// TIA Portal V20 export
// export: Created 2026-10-12T16:46:22.1158702Z, ExportSetting WithDefaults, DisplayName Totally Integrated Automation Portal, DisplayVersion V20 Update 6, DisplayName TIA Portal Openness, DisplayVersion V20 Update 6, DisplayName TIA Portal Version Control Interface, DisplayVersion V20 Update 6, DisplayName SINAMICS Startdrive Advanced, DisplayVersion V20 SP1 Update 2, DisplayName SINAMICS Startdrive G110M, G120, G120C, G120D, G120P, G115D, DisplayVersion V20 SP1 Update 2, DisplayName SINAMICS Startdrive G130, G150, S120, S150, SINAMICS MV, G220, S200, S210, DisplayVersion V20 SP1 Update 2, DisplayName STEP 7 Professional, DisplayVersion V20 Update 6, DisplayName STEP 7 Safety, DisplayVersion V20 Update 2, DisplayName WinCC Basic/Comfort/Advanced, DisplayVersion V20 Update 6, DisplayName WinCC Professional, DisplayVersion V20 Update 6, DisplayName WinCC Unified, DisplayVersion V20 Update 6
VAR_GLOBAL   // PLC tag table "Standard-Variablentabelle"
   "FI-Schutz 200F1 Heizung Bad 7 ist O.K." AT %I2.2 : Bool;
   "Sicherheitsschuetz Rueckfuehrung Heizung Bad 7" AT %I2.3 : Bool;
   "Heizung Bad 7 Keine uebertemperatur" AT %I2.4 : Bool;
   "Störmeldung Ultraschall Bad 7" AT %I2.6 : Bool;
   "Niveau Bad 7 OK" AT %I10.0 : Bool;
   "Pt100 Heizung Bad 7" AT %IW60 : Word;
   "FI-Schutz 210F1 Heizung Bad 8 ist O.K." AT %I2.7 : Bool;
   "Sicherheitsschuetz Rueckfuehrung Heizung Bad 8" AT %I3.0 : Bool;
   "Heizung Bad 8 Keine uebertemperatur" AT %I3.1 : Bool;
   "FILS Automat 213F1 Ultraschall Bad 8 ist O.K." AT %I3.2 : Bool;
   "Störmeldung Ultraschall Bad 8" AT %I3.3 : Bool;
   "Motorschutz 215Q1 Pumpe Bad 8 ist O.K." AT %I3.4 : Bool;
   "Wartungsschalter Pumpe Bad 8 ist eingeschaltet" AT %I3.5 : Bool;
   "Niveau Bad 8 OK" AT %I10.1 : Bool;
   "FI-Schutz 220F1 Heizung Bad 12 ist O.K." AT %I3.6 : Bool;
   "Sicherheitsschuetz Rueckfuehrung Heizung Bad 12" AT %I3.7 : Bool;
   "Heizung Bad 12 Keine uebertemperatur" AT %I4.0 : Bool;
   "FILS Automat 223F1 Ultraschall Bad 12 ist O.K." AT %I4.1 : Bool;
   "Störmeldung Ultraschall Bad 12" AT %I4.2 : Bool;
   "Motorschutz 225Q1 Pumpe Bad 12 ist O.K." AT %I4.3 : Bool;
   "Wartungsschalter Pumpe Bad 12 ist eingeschaltet" AT %I4.4 : Bool;
   "Niveau Bad 12 OK" AT %I10.2 : Bool;
   "Motorschutz 235Q1 Pumpe Bad 14 ist O.K." AT %I4.5 : Bool;
   "Wartungsschalter Pumpe Bad 14 ist eingeschaltet" AT %I4.6 : Bool;
   "Motorschutz 245Q1 Pumpe Bad 18 ist O.K." AT %I4.7 : Bool;
   "Wartungsschalter Pumpe Bad 18 ist eingeschaltet" AT %I5.0 : Bool;
   "Motorschutz 255Q1 Pumpe Bad 19 ist O.K." AT %I5.1 : Bool;
   "Wartungsschalter Pumpe Bad 19 ist eingeschaltet" AT %I5.2 : Bool;
   "Motorschutz 265Q1 Pumpe Bad 21 ist O.K." AT %I5.3 : Bool;
   "Wartungsschalter Pumpe Bad 21 ist eingeschaltet" AT %I5.4 : Bool;
   "Motorschutz und FI-Schutz 270Q1, 270F1 Heizung Bad 25 sind O.K." AT %I5.5 : Bool;
   "Motorschutz und FI-Schutz 271Q1, 271F1 Heizung Bad 25 sind O.K." AT %I5.6 : Bool;
   "Sicherheitsschuetze Rueckfuehrung Heizung Bad 25" AT %I5.7 : Bool;
   "Heizung Bad 25 Keine uebertemperatur" AT %I6.0 : Bool;
   "FILS Automat 274F1 Analysegerät Bad 25 ist O.K." AT %I6.1 : Bool;
   "Motorschutz 275Q1 Pumpe Bad 25 ist O.K." AT %I6.2 : Bool;
   "Wartungsschalter Pumpe Bad 25 ist eingeschaltet" AT %I6.3 : Bool;
   "Motorschutz 276Q1 Warenbewegung 1 Bad 25 ist O.K." AT %I6.4 : Bool;
   "Motorschutz 277Q1 Warenbewegung 2 Bad 25 ist O.K." AT %I6.5 : Bool;
   "FILS Automat 203F1 GR Wannenschutz Bad 25 ist O.K." AT %I2.5 : Bool;
   "Motorschutz 275aQ1 Pumpe Bad 25 ist O.K." AT %I8.7 : Bool;
   "Warenbewegung 1 Bad 25 FU bereit" AT %I9.5 : Bool;
   "Warenbewegung 2 Bad 25 FU bereit" AT %I9.6 : Bool;
   "Wartungsschalter Pumpe Bad 25 ist eingeschaltet(1)" AT %I9.7 : Bool;
   "Niveau Bad 25 OK" AT %I10.3 : Bool;
   "Motorschutz 285Q1 Pumpe Bad 26 ist O.K." AT %I6.6 : Bool;
   "Wartungsschalter Pumpe Bad 26 ist eingeschaltet" AT %I6.7 : Bool;
   "Motorschutz 295Q1 Pumpe Bad 31 ist O.K." AT %I7.0 : Bool;
   "Wartungsschalter Pumpe Bad 31 ist eingeschaltet" AT %I7.1 : Bool;
   "FI-Schutz 300F1 Heizung Bad 36 ist O.K." AT %I7.2 : Bool;
   "Sicherheitsschuetz Rueckfuehrung Heizung Bad 36" AT %I7.3 : Bool;
   "Heizung Bad 36 Keine uebertemperatur" AT %I7.4 : Bool;
   "Niveau Bad 36 OK" AT %I10.4 : Bool;
   "FI-Schutz 310F1 Heizung Bad 40 ist O.K." AT %I7.5 : Bool;
   "Sicherheitsschuetz Rueckfuehrung Heizung Bad 40" AT %I7.6 : Bool;
   "Heizung Bad 40 Keine uebertemperatur" AT %I7.7 : Bool;
   "Motorschutz 325Q1 Pumpe Bad 41 ist O.K." AT %I8.0 : Bool;
   "Wartungsschalter Pumpe Bad 41 ist eingeschaltet" AT %I8.1 : Bool;
   "Motorschutz 335Q1 Pumpe Bad 45 ist O.K." AT %I8.2 : Bool;
   "Wartungsschalter Pumpe Bad 45 ist eingeschaltet" AT %I8.3 : Bool;
   "FI-Schutz 340F1 Heizung Bad 46 ist O.K." AT %I8.4 : Bool;
   "Sicherheitsschuetz Rueckfuehrung Heizung Bad 46" AT %I8.5 : Bool;
   "Heizung Bad 46 Keine uebertemperatur" AT %I8.6 : Bool;
   "Niveau Bad 46 OK" AT %I10.6 : Bool;
   "Motorschutz 15Q0 Schaltschrankklimatisierung Feld 1-4 ist O.K." AT %I0.0 : Bool;
   "Klimagerät +E1-15A0 ist in Ordnung" AT %I0.1 : Bool;
   "Schaltschranktemperatur Feld 1 ist zu hoch" AT %I0.2 : Bool;
   "Schaltschranktemperatur Feld 2 ist zu hoch" AT %I0.3 : Bool;
   "FILS Automat 19F1 Schuko.Steckdosen PC-Bildschirm ist O.K." AT %I0.4 : Bool;
   "Not-Aus ist OK" AT %I0.5 : Bool;
   "Steuerspannung 31F1 Schaltschrank E1 ist O.K." AT %I1.0 : Bool;
   "Steuerspannung 31F3 SPS Out 1 ist O.K." AT %I1.1 : Bool;
   "Steuerspannung 31F5 SPS Out 2 ist O.K." AT %I1.2 : Bool;
   "Steuerspannung 31F6 SPS Out 3 ist O.K." AT %I1.3 : Bool;
   "Steuerspannung 31F8 Out 4 ist O.K." AT %I1.4 : Bool;
   "Steuerspannung 32F1 Rueckmeldung Wartungsschalter ist O.K." AT %I1.5 : Bool;
   "Steuerspannung 32F3 Sensorik 1 ist O.K." AT %I1.6 : Bool;
   "Busspannung 41F1 ist ok" AT %I1.7 : Bool;
   "Busspannung 41F2 ist ok" AT %I2.0 : Bool;
   "Busspannung 41F4 ist ok" AT %I2.1 : Bool;
   "Pt100 Heizung Bad 8" AT %IW62 : Word;
   "Pt100 Heizung Bad 12" AT %IW64 : Word;
   "Pt100 Heizung Bad 25" AT %IW66 : Word;
   "Pt100 Heizung Bad 36" AT %IW68 : Word;
   "Pt100 Heizung Bad 40" AT %IW70 : Word;
   "Pt100 Heizung Bad 46" AT %IW72 : Word;
   "FU Pumpe bereit" AT %I0.7 : Bool;
   Flexkraft_1 AT %IW500 : Word;
   Flexkraft_2 AT %IW502 : Word;
   Flexkraft_3 AT %IW504 : Word;
   Flexkraft_4 AT %IW506 : Word;
   Flexkraft_5 AT %IW508 : Word;
   Flexkraft_6 AT %IW510 : Word;
   Flexkraft_7 AT %IW512 : Word;
   Flexkraft_8 AT %IW514 : Word;
   Flexkraft_9 AT %IW516 : Word;
   Flexkraft_10 AT %IW518 : Word;
   "Niveau Bad 40 OK" AT %I10.5 : Bool;
   "Regelung Heizung Bad 7" AT %Q2.0 : Bool;
   "Sicherheitsschuetz Heizung Bad 7" AT %Q2.1 : Bool;
   "Pumpe Bad 8" AT %Q0.0 : Bool;
   "Regelung Heizung Bad 8" AT %Q2.2 : Bool;
   "Sicherheitsschuetz Heizung Bad 8" AT %Q2.3 : Bool;
   "Pumpe Bad 12" AT %Q0.1 : Bool;
   "Regelung Heizung Bad 12" AT %Q2.4 : Bool;
   "Sicherheitsschuetz Heizung Bad 12" AT %Q2.5 : Bool;
   "Pumpe Bad 14" AT %Q0.2 : Bool;
   "Pumpe Bad 18" AT %Q0.3 : Bool;
   "Pumpe Bad 19" AT %Q0.4 : Bool;
   "Pumpe Bad 21" AT %Q0.5 : Bool;
   "Netzschuetz Pumpe Bad 25" AT %Q0.6 : Bool;
   "Warenbewegung 1 Bad 25 Freigabe FU" AT %Q1.3 : Bool;
   "Warenbewegung 1 Bad 25 Reset FU" AT %Q1.4 : Bool;
   "Warenbewegung 2 Bad 25 Freigabe FU" AT %Q1.5 : Bool;
   "Warenbewegung 2 Bad 25 Reset FU" AT %Q1.6 : Bool;
   "Ansteuerung 275aK8" AT %Q1.7 : Bool;
   "Regelung Heizung 1 Bad 25" AT %Q2.6 : Bool;
   "Regelung Heizung 2 Bad 25" AT %Q2.7 : Bool;
   "Sicherheitsschuetze Heizung 1 + 2 Bad 25" AT %Q3.0 : Bool;
   "Warenbewegung 1 Bad 25 Netzschuetz" AT %Q3.1 : Bool;
   "Warenbewegung 2 Bad 25 Netzschuetz" AT %Q3.2 : Bool;
   "Pumpe Bad 26" AT %Q0.7 : Bool;
   "Pumpe Bad 31" AT %Q1.0 : Bool;
   "Regelung Heizung Bad 36" AT %Q3.3 : Bool;
   "Sicherheitsschuetz Heizung Bad 36" AT %Q3.4 : Bool;
   "Regelung Heizung Bad 40" AT %Q3.5 : Bool;
   "Sicherheitsschuetz Heizung Bad 40" AT %Q3.6 : Bool;
   "Pumpe Bad 41" AT %Q1.1 : Bool;
   "Pumpe Bad 45" AT %Q1.2 : Bool;
   "Regelung Heizung Bad 46" AT %Q3.7 : Bool;
   "Sicherheitsschuetz Heizung Bad 46" AT %Q4.0 : Bool;
   "Masch.Leuchte 1 Anlage Hupe" AT %Q4.1 : Bool;
   "Freigabe Ultraschall Pos. 8" AT %Q4.2 : Bool;
   "Freigabe Ultraschall Pos. 12" AT %Q4.3 : Bool;
   "Dosierpumpe 4 Ansteuerung" AT %Q4.4 : Bool;
   "Warenbewegung 1 Bad 25 Sollwert FU" AT %QW60 : Word;
   "Warenbewegung 2 Bad 25 Sollwert FU" AT %QW62 : Word;
   "Not-Aus Reset" AT %Q4.7 : Bool;
   Pumpen_FU_Steuerwert AT %QW64 : Word;
   "Reset FU Pumpe" AT %Q4.6 : Bool;
   "FU Pumpe Freigabe" AT %Q4.5 : Bool;
   System_Byte AT %MB1 : Byte;
   FirstScan AT %M1.0 : Bool;
   DiagStatusUpdate AT %M1.1 : Bool;
   AlwaysTRUE AT %M1.2 : Bool;
   AlwaysFALSE AT %M1.3 : Bool;
   Clock_Byte AT %MB0 : Byte;
   Clock_10Hz AT %M0.0 : Bool;
   Clock_5Hz AT %M0.1 : Bool;
   "Clock_2.5Hz" AT %M0.2 : Bool;
   Clock_2Hz AT %M0.3 : Bool;
   "Clock_1.25Hz" AT %M0.4 : Bool;
   Clock_1Hz AT %M0.5 : Bool;
   "Clock_0.625Hz" AT %M0.6 : Bool;
   "Clock_0.5Hz" AT %M0.7 : Bool;
   User_Level AT %MW10 : Int;   // User Level von aktiven User
   Empty AT %M100.0 : Bool;
   Empty1 AT %MW101 : Int;
   Flexkraft_11 AT %QW500 : Word;
   Flexkraft_12 AT %QW502 : Word;
   Flexkraft_13 AT %QW504 : Word;
   Flexkraft_14 AT %QW506 : Word;
   Flexkraft_15 AT %QW508 : Word;
   Flexkraft_16 AT %QW510 : Word;
   Flexkraft_17 AT %QW512 : Word;
   Flexkraft_18 AT %QW514 : Word;
   Flexkraft_19 AT %QW516 : Word;
   Flexkraft_20 AT %IW532 : Word;
   Flexkraft_21 AT %IW534 : Word;
   Flexkraft_22 AT %IW536 : Word;
   Flexkraft_23 AT %IW538 : Word;
   Flexkraft_24 AT %IW540 : Word;
   Flexkraft_25 AT %IW542 : Word;
   Flexkraft_26 AT %IW544 : Word;
   Flexkraft_27 AT %IW546 : Word;
   Flexkraft_28 AT %IW548 : Word;
   Flexkraft_29 AT %IW550 : Word;
   Flexkraft_30 AT %IW564 : Word;
   Flexkraft_31 AT %IW566 : Word;
   Flexkraft_32 AT %IW568 : Word;
   Flexkraft_33 AT %IW570 : Word;
   Flexkraft_34 AT %IW572 : Word;
   Flexkraft_35 AT %IW574 : Word;
   Flexkraft_36 AT %IW576 : Word;
   Flexkraft_37 AT %IW578 : Word;
   Flexkraft_38 AT %IW580 : Word;
   Flexkraft_39 AT %IW582 : Word;
   Flexkraft_40 AT %QW532 : Word;
   Flexkraft_41 AT %QW534 : Word;
   Flexkraft_42 AT %QW536 : Word;
   Flexkraft_43 AT %QW538 : Word;
   Flexkraft_44 AT %QW540 : Word;
   Flexkraft_45 AT %QW542 : Word;
   Flexkraft_46 AT %QW544 : Word;
   Flexkraft_47 AT %QW564 : Word;
   Flexkraft_48 AT %QW548 : Word;
   Flexkraft_49 AT %QW546 : Word;
   Flexkraft_50 AT %QW566 : Word;
   Flexkraft_51 AT %QW568 : Word;
   Flexkraft_52 AT %QW570 : Word;
   Flexkraft_53 AT %QW574 : Word;
   Flexkraft_54 AT %QW572 : Word;
   Flexkraft_55 AT %QW576 : Word;
   Flexkraft_56 AT %QW578 : Word;
   Flexkraft_57 AT %QW580 : Word;
   "Alarm Walchem Controller" AT %I0.6 : Bool;
END_VAR
VAR_GLOBAL CONSTANT   // user constants
   c_Prozessgruppen : Int := 6;
   c_Anzahl_Benutzer : Int := 20;
   c_Anzahl_Artikel : Int := 50;
   c_Anzahl_Bad : Int := 47;
END_VAR
